FUNCTION F_WordToRange : REAL
VAR_INPUT
	wWord 					:WORD;
	rLowLimit 				:REAL;
	rHighLimit 				:REAL;
END_VAR
VAR
END_VAR


F_WordToRange := (rHighLimit - rLowLimit) * WORD_TO_REAL(wWord) * 0.00001525902189669640 + rLowLimit;

END_FUNCTION

(* stored: Version 1.1.0.1, ProductVersion 3.1.4024.15
   POU F_WordToRange: Id {eff690ad-d198-4dfc-94cd-00264b5c1195}, SpecialFunc None *)
